Fanuc KAREL source: KT00584.KL

PROGRAM KT00584
%NOLOCKGROUP
VAR
  I1: INTEGER
  V2: VECTOR
  OUT: VECTOR
BEGIN
  I1 = 2
    V2.Y = 2.0
  OUT = I1 - V2
END KT00584
